Fanuc KAREL source: KD00009.KL

PROGRAM KD00009
%NOLOCKGROUP
%DELAY = 100
VAR
  I: INTEGER
  J: INTEGER
  B: BOOLEAN
  R: REAL
  S: STRING[80]
BEGIN
  I = 1
END KD00009
